// Objet qui réagit au changement d'OF (compteur, P3 : remise à zéro au changement d'OF, docs/03 § 8.4)
INTERFACE I_OrderAware

METHOD OnOrderChange
END_METHOD

END_INTERFACE

(* stored: Version 1.1.0.1, ProductVersion 3.1.4024.12
   Itf I_OrderAware: Id {5e10a71e-c4e1-5cb0-a931-39a1214c6a5f}
   Method OnOrderChange: Id {ecd8779a-a207-5565-a570-fe6ef8cc88dc} *)
